Fanuc KAREL source: kd00033.KL

-- PROVISIONAL review KL for V940-1; original PC SHA256 97f157aa6b4e6439c3d189a54e428837f283c6c7727d4f34ee29fdb45ccf6144
-- Incomplete behavior may be omitted. Consult companion uncertainty JSON. Do not deploy.
PROGRAM KD00033
%NOLOCKGROUP
VAR
  I : INTEGER
  J : INTEGER
  B : BOOLEAN
  R : REAL
  S : STRING[80]
BEGIN
  -- V9_ZERO_TABLE_METADATA_HINT layout=0001; no indexed target words; source/name/runtime held
  -- UNRESOLVED_PC offsets 5-24; opcodes 9D,81,18,9D,1B,9D,12,22,9D,13,04
  -- UNRESOLVED_PC offsets 29-33; opcodes 7F
END KD00033
